FUNCTION_BLOCK SortingCycleCoordinator (* Minimal Reset, Run and Stop controller. Standard equipment and movement sequences remain separate. *)
  (* Standard: 61499-2 *)
  (* Version 2.0, 2026-11-09, sorting2n, sorting2n *)
  PACKAGE Main;
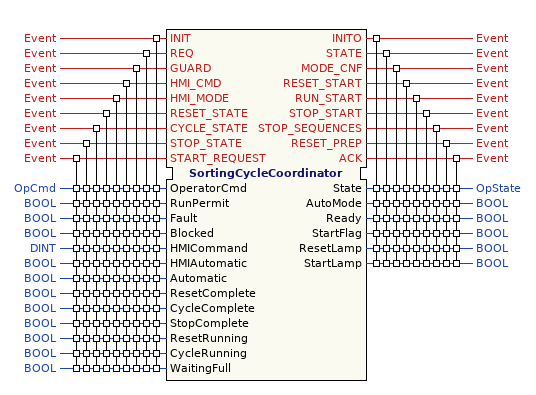
  EVENT_INPUT
    INIT WITH OperatorCmd, RunPermit, Fault, Blocked, HMICommand, HMIAutomatic, Automatic, ResetComplete, CycleComplete, StopComplete, ResetRunning, CycleRunning, WaitingFull;
    REQ WITH OperatorCmd, RunPermit, Fault, Blocked, HMICommand, HMIAutomatic, Automatic, ResetComplete, CycleComplete, StopComplete, ResetRunning, CycleRunning, WaitingFull;
    GUARD WITH OperatorCmd, RunPermit, Fault, Blocked, HMICommand, HMIAutomatic, Automatic, ResetComplete, CycleComplete, StopComplete, ResetRunning, CycleRunning, WaitingFull;
    HMI_CMD WITH OperatorCmd, RunPermit, Fault, Blocked, HMICommand, HMIAutomatic, Automatic, ResetComplete, CycleComplete, StopComplete, ResetRunning, CycleRunning, WaitingFull;
    HMI_MODE WITH OperatorCmd, RunPermit, Fault, Blocked, HMICommand, HMIAutomatic, Automatic, ResetComplete, CycleComplete, StopComplete, ResetRunning, CycleRunning, WaitingFull;
    RESET_STATE WITH OperatorCmd, RunPermit, Fault, Blocked, HMICommand, HMIAutomatic, Automatic, ResetComplete, CycleComplete, StopComplete, ResetRunning, CycleRunning, WaitingFull;
    CYCLE_STATE WITH OperatorCmd, RunPermit, Fault, Blocked, HMICommand, HMIAutomatic, Automatic, ResetComplete, CycleComplete, StopComplete, ResetRunning, CycleRunning, WaitingFull;
    STOP_STATE WITH OperatorCmd, RunPermit, Fault, Blocked, HMICommand, HMIAutomatic, Automatic, ResetComplete, CycleComplete, StopComplete, ResetRunning, CycleRunning, WaitingFull;
    START_REQUEST WITH OperatorCmd, RunPermit, Fault, Blocked, HMICommand, HMIAutomatic, Automatic, ResetComplete, CycleComplete, StopComplete, ResetRunning, CycleRunning, WaitingFull;
  END_EVENT
  EVENT_OUTPUT
    INITO WITH State, AutoMode, Ready, StartFlag, ResetLamp, StartLamp;
    STATE WITH State, AutoMode, Ready, StartFlag, ResetLamp, StartLamp;
    MODE_CNF WITH State, AutoMode, Ready, StartFlag, ResetLamp, StartLamp;
    RESET_START WITH State, AutoMode, Ready, StartFlag, ResetLamp, StartLamp;
    RUN_START WITH State, AutoMode, Ready, StartFlag, ResetLamp, StartLamp;
    STOP_START WITH State, AutoMode, Ready, StartFlag, ResetLamp, StartLamp;
    STOP_SEQUENCES WITH State, AutoMode, Ready, StartFlag, ResetLamp, StartLamp;
    RESET_PREP WITH State, AutoMode, Ready, StartFlag, ResetLamp, StartLamp;
    ACK WITH State, AutoMode, Ready, StartFlag, ResetLamp, StartLamp;
  END_EVENT
  VAR_INPUT
    OperatorCmd : OpCmd;
    RunPermit : BOOL;
    Fault : BOOL;
    Blocked : BOOL;
    HMICommand : DINT;
    HMIAutomatic : BOOL;
    Automatic : BOOL;
    ResetComplete : BOOL;
    CycleComplete : BOOL;
    StopComplete : BOOL;
    ResetRunning : BOOL := FALSE;
    CycleRunning : BOOL := FALSE;
    WaitingFull : BOOL := FALSE;
  END_VAR
  VAR_OUTPUT
    State : OpState;
    AutoMode : BOOL := FALSE;
    Ready : BOOL := FALSE;
    StartFlag : BOOL := FALSE;
    ResetLamp : BOOL := FALSE;
    StartLamp : BOOL := FALSE;
  END_VAR
  VAR
    Action : DINT;
    Requested : DINT;
  END_VAR
  EC_STATES
    IDLE;
    INITIALIZE : INITIALIZE, NOP -> STOP_SEQUENCES, NOP -> STATE, NOP -> INITO;
    ON_REQ : ON_REQ;
    ON_HMI_CMD : ON_HMI_CMD;
    ON_GUARD : ON_GUARD;
    ON_RESET_STATE : ON_RESET_STATE;
    ON_CYCLE_STATE : ON_CYCLE_STATE;
    ON_STOP_STATE : ON_STOP_STATE;
    SET_MODE : SET_MODE, NOP -> MODE_CNF;
    RESET : RESET, NOP -> STOP_SEQUENCES, NOP -> RESET_PREP, NOP -> STATE, NOP -> RESET_START;
    RUN : RUN, NOP -> STOP_SEQUENCES, NOP -> STATE, NOP -> RUN_START;
    STOP : STOP, NOP -> STOP_SEQUENCES, NOP -> STATE, NOP -> STOP_START;
    RESET_DONE : RESET_DONE, NOP -> STATE;
    RUN_DONE : RUN_DONE, NOP -> STATE;
    STOP_DONE : STOP_DONE, NOP -> STATE;
    RESET_OBSERVED : RESET_OBSERVED, NOP -> STATE;
    RUN_OBSERVED : RUN_OBSERVED, NOP -> STATE;
    ACKNOWLEDGE : ACKNOWLEDGE, NOP -> ACK;
    ON_START_REQUEST : ON_START_REQUEST;
  END_STATES
  EC_TRANSITIONS
    IDLE TO INITIALIZE := INIT;
    INITIALIZE TO IDLE := 1;
    IDLE TO ON_REQ := REQ;
    ON_REQ TO RESET := Action = 1;
    ON_REQ TO RUN := Action = 2;
    ON_REQ TO STOP := Action = 3;
    ON_REQ TO RESET_DONE := Action = 4;
    ON_REQ TO RUN_DONE := Action = 5;
    ON_REQ TO STOP_DONE := Action = 6;
    ON_REQ TO RESET_OBSERVED := Action = 7;
    ON_REQ TO RUN_OBSERVED := Action = 8;
    ON_REQ TO ACKNOWLEDGE := Action = 9;
    ON_REQ TO IDLE := 1;
    IDLE TO ON_HMI_CMD := HMI_CMD;
    ON_HMI_CMD TO RESET := Action = 1;
    ON_HMI_CMD TO RUN := Action = 2;
    ON_HMI_CMD TO STOP := Action = 3;
    ON_HMI_CMD TO RESET_DONE := Action = 4;
    ON_HMI_CMD TO RUN_DONE := Action = 5;
    ON_HMI_CMD TO STOP_DONE := Action = 6;
    ON_HMI_CMD TO RESET_OBSERVED := Action = 7;
    ON_HMI_CMD TO RUN_OBSERVED := Action = 8;
    ON_HMI_CMD TO ACKNOWLEDGE := Action = 9;
    ON_HMI_CMD TO IDLE := 1;
    IDLE TO ON_GUARD := GUARD;
    ON_GUARD TO RESET := Action = 1;
    ON_GUARD TO RUN := Action = 2;
    ON_GUARD TO STOP := Action = 3;
    ON_GUARD TO RESET_DONE := Action = 4;
    ON_GUARD TO RUN_DONE := Action = 5;
    ON_GUARD TO STOP_DONE := Action = 6;
    ON_GUARD TO RESET_OBSERVED := Action = 7;
    ON_GUARD TO RUN_OBSERVED := Action = 8;
    ON_GUARD TO ACKNOWLEDGE := Action = 9;
    ON_GUARD TO IDLE := 1;
    IDLE TO ON_RESET_STATE := RESET_STATE;
    ON_RESET_STATE TO RESET := Action = 1;
    ON_RESET_STATE TO RUN := Action = 2;
    ON_RESET_STATE TO STOP := Action = 3;
    ON_RESET_STATE TO RESET_DONE := Action = 4;
    ON_RESET_STATE TO RUN_DONE := Action = 5;
    ON_RESET_STATE TO STOP_DONE := Action = 6;
    ON_RESET_STATE TO RESET_OBSERVED := Action = 7;
    ON_RESET_STATE TO RUN_OBSERVED := Action = 8;
    ON_RESET_STATE TO ACKNOWLEDGE := Action = 9;
    ON_RESET_STATE TO IDLE := 1;
    IDLE TO ON_CYCLE_STATE := CYCLE_STATE;
    ON_CYCLE_STATE TO RESET := Action = 1;
    ON_CYCLE_STATE TO RUN := Action = 2;
    ON_CYCLE_STATE TO STOP := Action = 3;
    ON_CYCLE_STATE TO RESET_DONE := Action = 4;
    ON_CYCLE_STATE TO RUN_DONE := Action = 5;
    ON_CYCLE_STATE TO STOP_DONE := Action = 6;
    ON_CYCLE_STATE TO RESET_OBSERVED := Action = 7;
    ON_CYCLE_STATE TO RUN_OBSERVED := Action = 8;
    ON_CYCLE_STATE TO ACKNOWLEDGE := Action = 9;
    ON_CYCLE_STATE TO IDLE := 1;
    IDLE TO ON_STOP_STATE := STOP_STATE;
    ON_STOP_STATE TO RESET := Action = 1;
    ON_STOP_STATE TO RUN := Action = 2;
    ON_STOP_STATE TO STOP := Action = 3;
    ON_STOP_STATE TO RESET_DONE := Action = 4;
    ON_STOP_STATE TO RUN_DONE := Action = 5;
    ON_STOP_STATE TO STOP_DONE := Action = 6;
    ON_STOP_STATE TO RESET_OBSERVED := Action = 7;
    ON_STOP_STATE TO RUN_OBSERVED := Action = 8;
    ON_STOP_STATE TO ACKNOWLEDGE := Action = 9;
    ON_STOP_STATE TO IDLE := 1;
    IDLE TO SET_MODE := HMI_MODE;
    SET_MODE TO IDLE := 1;
    RESET TO IDLE := 1;
    RUN TO IDLE := 1;
    STOP TO IDLE := 1;
    RESET_DONE TO IDLE := 1;
    RUN_DONE TO IDLE := 1;
    STOP_DONE TO IDLE := 1;
    RESET_OBSERVED TO IDLE := 1;
    RUN_OBSERVED TO IDLE := 1;
    ACKNOWLEDGE TO IDLE := 1;
    IDLE TO ON_START_REQUEST := START_REQUEST;
    ON_START_REQUEST TO RESET := Action = 1;
    ON_START_REQUEST TO RUN := Action = 2;
    ON_START_REQUEST TO STOP := Action = 3;
    ON_START_REQUEST TO RESET_DONE := Action = 4;
    ON_START_REQUEST TO RUN_DONE := Action = 5;
    ON_START_REQUEST TO STOP_DONE := Action = 6;
    ON_START_REQUEST TO RESET_OBSERVED := Action = 7;
    ON_START_REQUEST TO RUN_OBSERVED := Action = 8;
    ON_START_REQUEST TO ACKNOWLEDGE := Action = 9;
    ON_START_REQUEST TO IDLE := 1;
  END_TRANSITIONS
  ALGORITHM INITIALIZE IN ST:
State := SE.App2StateManagement.OpState#PhaseStopped; Ready := FALSE; AutoMode := Automatic; Action := 0; Requested := 0;

StartFlag := FALSE; StartLamp := FALSE; ResetLamp := TRUE;
  END_ALGORITHM
  ALGORITHM ON_REQ IN ST:
Requested := OperatorCmd;
Action := 0;
IF Requested = 2 AND WaitingFull AND State = SE.App2StateManagement.OpState#PhaseExecute THEN Action := 9;
ELSIF Requested = 3 OR Requested = 4 OR Requested = 6 OR Requested = 8 THEN IF State <> SE.App2StateManagement.OpState#PhaseStopping THEN Action := 3; END_IF;
ELSIF Requested = 1 AND RunPermit THEN IF State = SE.App2StateManagement.OpState#PhaseStopped OR State = SE.App2StateManagement.OpState#PhaseIdle THEN Action := 1; END_IF;
ELSIF Requested = 2 AND Ready AND RunPermit AND NOT Fault AND State = SE.App2StateManagement.OpState#PhaseIdle THEN Action := 2;
END_IF;
  END_ALGORITHM
  ALGORITHM ON_HMI_CMD IN ST:
Requested := HMICommand;
Action := 0;
IF Requested = 2 AND WaitingFull AND State = SE.App2StateManagement.OpState#PhaseExecute THEN Action := 9;
ELSIF Requested = 3 OR Requested = 4 OR Requested = 6 OR Requested = 8 THEN IF State <> SE.App2StateManagement.OpState#PhaseStopping THEN Action := 3; END_IF;
ELSIF Requested = 1 AND RunPermit THEN IF State = SE.App2StateManagement.OpState#PhaseStopped OR State = SE.App2StateManagement.OpState#PhaseIdle THEN Action := 1; END_IF;
ELSIF Requested = 2 AND Ready AND RunPermit AND NOT Fault AND State = SE.App2StateManagement.OpState#PhaseIdle THEN Action := 2;
END_IF;
  END_ALGORITHM
  ALGORITHM ON_GUARD IN ST:
Action := 0;
StartLamp := (State = SE.App2StateManagement.OpState#PhaseIdle) OR WaitingFull;
ResetLamp := (State = SE.App2StateManagement.OpState#PhaseStopped) AND NOT Ready;
IF (State = SE.App2StateManagement.OpState#PhaseExecute OR State = SE.App2StateManagement.OpState#PhaseResetting) AND (NOT RunPermit OR Fault) THEN Action := 3; END_IF;
  END_ALGORITHM
  ALGORITHM ON_RESET_STATE IN ST:
Action := 0;
IF ResetComplete AND State = SE.App2StateManagement.OpState#PhaseResetting THEN Action := 4;
ELSIF ResetRunning AND State <> SE.App2StateManagement.OpState#PhaseResetting AND State <> SE.App2StateManagement.OpState#PhaseStopping THEN Action := 7; END_IF;
  END_ALGORITHM
  ALGORITHM ON_CYCLE_STATE IN ST:
Action := 0;
IF CycleComplete AND State = SE.App2StateManagement.OpState#PhaseExecute THEN Action := 5;
ELSIF CycleRunning AND Ready AND RunPermit AND NOT Fault AND State = SE.App2StateManagement.OpState#PhaseIdle THEN Action := 8; END_IF;
  END_ALGORITHM
  ALGORITHM ON_STOP_STATE IN ST:
Action := 0; IF StopComplete AND State = SE.App2StateManagement.OpState#PhaseStopping THEN Action := 6; END_IF;
  END_ALGORITHM
  ALGORITHM SET_MODE IN ST:
AutoMode := HMIAutomatic;
  END_ALGORITHM
  ALGORITHM RESET IN ST:
State := SE.App2StateManagement.OpState#PhaseResetting; Ready := FALSE;

StartFlag := FALSE; StartLamp := FALSE; ResetLamp := FALSE;
  END_ALGORITHM
  ALGORITHM RUN IN ST:
State := SE.App2StateManagement.OpState#PhaseExecute;

StartFlag := TRUE; StartLamp := FALSE; ResetLamp := FALSE;
  END_ALGORITHM
  ALGORITHM STOP IN ST:
State := SE.App2StateManagement.OpState#PhaseStopping; Ready := FALSE;

StartFlag := FALSE; StartLamp := FALSE; ResetLamp := TRUE;
  END_ALGORITHM
  ALGORITHM RESET_DONE IN ST:
State := SE.App2StateManagement.OpState#PhaseIdle; Ready := TRUE;

StartFlag := FALSE; StartLamp := TRUE; ResetLamp := FALSE;
  END_ALGORITHM
  ALGORITHM RUN_DONE IN ST:
State := SE.App2StateManagement.OpState#PhaseIdle; Ready := TRUE;

StartFlag := FALSE; StartLamp := TRUE; ResetLamp := FALSE;
  END_ALGORITHM
  ALGORITHM STOP_DONE IN ST:
State := SE.App2StateManagement.OpState#PhaseStopped; Ready := FALSE;

StartFlag := FALSE; StartLamp := FALSE; ResetLamp := TRUE;
  END_ALGORITHM
  ALGORITHM NOP IN ST:
Action := Action;
  END_ALGORITHM
  ALGORITHM RESET_OBSERVED IN ST:
State := SE.App2StateManagement.OpState#PhaseResetting; Ready := FALSE; StartFlag := FALSE; ResetLamp := FALSE; StartLamp := FALSE;
  END_ALGORITHM
  ALGORITHM RUN_OBSERVED IN ST:
State := SE.App2StateManagement.OpState#PhaseExecute; StartFlag := TRUE; StartLamp := FALSE; ResetLamp := FALSE;
  END_ALGORITHM
  ALGORITHM ACKNOWLEDGE IN ST:
Action := 0;
  END_ALGORITHM
  ALGORITHM ON_START_REQUEST IN ST:
Requested := 2;
Action := 0;
IF Requested = 2 AND WaitingFull AND State = SE.App2StateManagement.OpState#PhaseExecute THEN Action := 9;
ELSIF Requested = 3 OR Requested = 4 OR Requested = 6 OR Requested = 8 THEN IF State <> SE.App2StateManagement.OpState#PhaseStopping THEN Action := 3; END_IF;
ELSIF Requested = 1 AND RunPermit THEN IF State = SE.App2StateManagement.OpState#PhaseStopped OR State = SE.App2StateManagement.OpState#PhaseIdle THEN Action := 1; END_IF;
ELSIF Requested = 2 AND Ready AND RunPermit AND NOT Fault AND State = SE.App2StateManagement.OpState#PhaseIdle THEN Action := 2;
END_IF;
  END_ALGORITHM
END_FUNCTION_BLOCK
